Fanuc KAREL source: KT00893.KL

PROGRAM KT00893
%NOLOCKGROUP
VAR
  P1: POSITION
  P2: POSITION
  OUT: BOOLEAN
BEGIN
  OUT = IN_RANGE(P1)
END KT00893
